Fanuc KAREL source: KA00163.KL

PROGRAM KA00163
%NOLOCKGROUP
VAR
  SRC: ARRAY[4] OF BOOLEAN
  DST: ARRAY[4] OF INTEGER
BEGIN
  DST = SRC
END KA00163
